(* IEC 61131-3 sources: trust-platform/examples/control/03-production-quality-digital-pid/38-positional-incremental-pid/src, 2 files *)

(* ---- Main.st ---- *)
USING Control;

(* Fraction of the raw-minus-filtered difference applied per update: alpha = dt/(Tf + dt). *)
FUNCTION FilterFraction : LREAL
VAR_INPUT
    CycleTime : LREAL;
    FilterTime : LREAL;
END_VAR
FilterFraction := CycleTime / (FilterTime + CycleTime);
END_FUNCTION

(* One first-order filter update: the filtered value moves alpha of the way toward the raw value. *)
FUNCTION FilterUpdate : LREAL
VAR_INPUT
    PreviousFilteredValue : LREAL;
    RawValue : LREAL;
    FilterFraction : LREAL;
END_VAR
FilterUpdate := PreviousFilteredValue + FilterFraction * (RawValue - PreviousFilteredValue);
END_FUNCTION

FUNCTION SamePidParameters : BOOL
VAR_INPUT
    Left : Control.PIDParameters;
    Right : Control.PIDParameters;
END_VAR
SamePidParameters :=
    Left.ProportionalGain = Right.ProportionalGain
    AND Left.IntegralGain = Right.IntegralGain
    AND Left.DerivativeGain = Right.DerivativeGain
    AND Left.ProportionalSetpointWeight = Right.ProportionalSetpointWeight
    AND Left.DerivativeSetpointWeight = Right.DerivativeSetpointWeight
    AND Left.Bias = Right.Bias
    AND Left.OutputMinimum = Right.OutputMinimum
    AND Left.OutputMaximum = Right.OutputMaximum
    AND Left.RateMinimum = Right.RateMinimum
    AND Left.RateMaximum = Right.RateMaximum
    AND Left.TrackingTime = Right.TrackingTime
    AND Left.AntiWindup = Right.AntiWindup;
END_FUNCTION

(* The positional form of this lesson's PID (β = 1, γ = 0): the complete request every update, from its own
   retained integral. Three rules make it the same controller as the incremental form of Control.PID:
   tracking corrects the integral after the clamp, in Manual the integral follows the manual torque, and a
   gain revision moves the change of the previous P and D into the integral. *)
FUNCTION_BLOCK PositionalPid
VAR_INPUT
    Parameters : Control.PIDParameters;
    Input : Control.PIDInput;
    PreloadOnGainRevision : BOOL := TRUE;
END_VAR
VAR_OUTPUT
    ErrorRad : LREAL;
    ProportionalNm : LREAL;
    TrialIntegralNm : LREAL;
    DerivativeNm : LREAL;
    RequestNm : LREAL;
    TorqueNm : LREAL;
    IntegralNm : LREAL;
END_VAR
VAR
    ProportionalGain : LREAL;
    DerivativeGain : LREAL;
    VelocityRadS : LREAL;
    PreviousAngleRad : LREAL;
    PreviousErrorRad : LREAL;
    PreviousVelocityRadS : LREAL;
END_VAR
(* Gain revision: P and D of the previous update change by (Kp,old − Kp,new)·e and (Kd,new − Kd,old)·ω_f;
   the integral takes that over, so the retained request stays the same. *)
IF PreloadOnGainRevision THEN
    IntegralNm := IntegralNm
        + (ProportionalGain - Parameters.ProportionalGain) * PreviousErrorRad
        - (DerivativeGain - Parameters.DerivativeGain) * PreviousVelocityRadS;
END_IF;
ProportionalGain := Parameters.ProportionalGain;
DerivativeGain := Parameters.DerivativeGain;

ErrorRad := Input.Setpoint - Input.ProcessValue;
VelocityRadS := (Input.ProcessValue - PreviousAngleRad) / Input.CycleTime;
ProportionalNm := ProportionalGain * ErrorRad;
DerivativeNm := -DerivativeGain * VelocityRadS;
IF Input.Mode = PIDMode#Auto THEN
    TrialIntegralNm := IntegralNm + Parameters.IntegralGain * ErrorRad * Input.CycleTime;
    RequestNm := ProportionalNm + TrialIntegralNm + DerivativeNm;
    TorqueNm := LIMIT(Parameters.OutputMinimum, RequestNm, Parameters.OutputMaximum);
    IntegralNm := TrialIntegralNm + Input.CycleTime / Parameters.TrackingTime * (TorqueNm - RequestNm);
ELSE
    (* Manual: the integral follows the manual torque, so the first Auto update continues from it. *)
    RequestNm := Input.ManualOutput;
    TorqueNm := LIMIT(Parameters.OutputMinimum, Input.ManualOutput, Parameters.OutputMaximum);
    IntegralNm := Input.ManualOutput - ProportionalNm - DerivativeNm;
    TrialIntegralNm := IntegralNm;
END_IF;
PreviousAngleRad := Input.ProcessValue;
PreviousErrorRad := ErrorRad;
PreviousVelocityRadS := VelocityRadS;
END_FUNCTION_BLOCK

PROGRAM Main
VAR
    Controller : Control.PID;
    (* The discrete PID of Lesson 38: Kp = 16 N·m/rad, Ki = 4 N·m/(rad·s), Kd = 7 N·m·s/rad on the
       filtered angle, the full target change in P, ±20 N·m with back-calculation (Tt = 1 s). *)
    Parameters : Control.PIDParameters := (
        ProportionalGain := LREAL#16.0,
        IntegralGain := LREAL#4.0,
        DerivativeGain := LREAL#7.0,
        ProportionalSetpointWeight := LREAL#1.0,
        DerivativeSetpointWeight := LREAL#0.0,
        Bias := LREAL#0.0,
        OutputMinimum := LREAL#-20.0,
        OutputMaximum := LREAL#20.0,
        RateMinimum := LREAL#-10000.0,
        RateMaximum := LREAL#10000.0,
        TrackingTime := LREAL#1.0,
        AntiWindup := PIDAntiWindup#BackCalculation
    );
    ConfiguredParameters : Control.PIDParameters;
    ParameterRevision : DINT := 0;
    InitialState : Control.PIDInitialState;
    Input : Control.PIDInput;
    Initialized : BOOL := FALSE;
    AutoMode : BOOL := FALSE;
    ManualTorqueNm : LREAL := 0.0;
    SafetyAbort : BOOL := FALSE;
    SetpointRad : LREAL := 0.0;
    AngleRad : LREAL := 0.0;
    VelocityRadS : LREAL := 0.0;
    TorqueNm : LREAL := 0.0;
    (* Drum load of the simulated test rig, in N·m: the experiment couples a 2 kg weight at the 0.1 m drum
       radius, 1.962 N·m. The controller does not use it. *)
    LoadTorqueNm : LREAL := 0.0;
    (* Measurement filter on the angle: Control.PID differentiates the filtered angle, so D uses the
       filtered velocity. Tf = 0 bypasses the filter. *)
    FilterTimeS : LREAL := 0.1;
    FilterAlpha : LREAL := 1.0;
    FilteredAngleRad : LREAL := 0.0;
    FilterActive : BOOL := FALSE;
    FilterWasActive : BOOL := FALSE;
    (* Three other forms, each updated from the same Input as Controller. None of them drives the axis. *)
    Positional : PositionalPid;
    Unpreloaded : PositionalPid;
    RetainedApplied : Control.PID;
    RetainedAppliedParameters : Control.PIDParameters;
    PositionalTorqueNm : LREAL := 0.0;
    UnpreloadedTorqueNm : LREAL := 0.0;
    RetainedAppliedTorqueNm : LREAL := 0.0;
    ErrorRad : LREAL := 0.0;
    ProportionalNm : LREAL := 0.0;
    DerivativeNm : LREAL := 0.0;
    RequestNm : LREAL := 0.0;
    IntegralNm : LREAL := 0.0;
    (* Project experiment. *)
    ExperimentEnabled : BOOL := FALSE;
    ExperimentWasEnabled : BOOL := FALSE;
    Active : BOOL := FALSE;
    ExperimentUpdates : DINT := 0;
    GainBeforeRevision : LREAL := 16.0;
    (* Software travel and speed limits of the axis. *)
    AngleLimitRad : LREAL := 2.0;
    VelocityLimitRadS : LREAL := 10.0;
END_VAR

(* Leaving the travel or speed range removes the torque until a full restart. *)
IF ABS(AngleRad) > AngleLimitRad OR ABS(VelocityRadS) > VelocityLimitRadS THEN
    SafetyAbort := TRUE;
END_IF;

(* Control Studio's project experiment couples the drum load and steps the target to 1.5 rad in Auto; 1 s
   later it applies Kp = 24 N·m/rad, as a gain revision would. Its end uncouples the load, restores the gain
   and returns to Manual with zero torque. *)
IF ExperimentEnabled AND NOT ExperimentWasEnabled THEN
    Active := TRUE;
    ExperimentUpdates := 0;
    LoadTorqueNm := LREAL#1.962;
    SetpointRad := LREAL#1.5;
    AutoMode := TRUE;
ELSIF NOT ExperimentEnabled AND ExperimentWasEnabled THEN
    Active := FALSE;
    LoadTorqueNm := LREAL#0.0;
    AutoMode := FALSE;
    SetpointRad := AngleRad;
    IF ExperimentUpdates > 50 THEN
        Parameters.ProportionalGain := GainBeforeRevision;
    END_IF;
END_IF;
ExperimentWasEnabled := ExperimentEnabled;
IF Active THEN
    IF ExperimentUpdates = 50 THEN
        GainBeforeRevision := Parameters.ProportionalGain;
        Parameters.ProportionalGain := LREAL#24.0;
    END_IF;
    ExperimentUpdates := ExperimentUpdates + 1;
END_IF;

(* Control Studio's Apply replaces this complete record at the task boundary. *)
IF NOT Initialized OR NOT SamePidParameters(Left := Parameters, Right := ConfiguredParameters) THEN
    ConfiguredParameters := Parameters;
    ParameterRevision := ParameterRevision + 1;
END_IF;
Controller.Configure(Parameters := Parameters);
(* Tracking with Tt = Δt removes the whole excess: this controller retains the applied torque. *)
RetainedAppliedParameters := Parameters;
RetainedAppliedParameters.TrackingTime := LREAL#0.02;
RetainedApplied.Configure(Parameters := RetainedAppliedParameters);

IF NOT Initialized THEN
    (* Hot reset: the axis rests without torque and the setpoint follows the measured angle. *)
    ManualTorqueNm := LREAL#0.0;
    IF NOT AutoMode THEN
        SetpointRad := AngleRad;
    END_IF;
    InitialState.Setpoint := SetpointRad;
    InitialState.ProcessValue := AngleRad;
    InitialState.NominalOutput := ManualTorqueNm;
    InitialState.SaturatedOutput := ManualTorqueNm;
    InitialState.SetpointRate := LREAL#0.0;
    InitialState.ProcessValueRate := LREAL#0.0;
    InitialState.FeedForward := LREAL#0.0;
    Controller.Initialize(State := InitialState);
    RetainedApplied.Initialize(State := InitialState);
    Initialized := TRUE;
END_IF;

(* The filter runs while the controller is in Auto. In Manual and in the Auto-entry scan it restarts
   from the measurement, so entering Auto is exactly bumpless; filtering starts with the next scan. *)
FilterAlpha := FilterFraction(CycleTime := LREAL#0.02, FilterTime := MAX(FilterTimeS, LREAL#0.0));
FilterActive := AutoMode AND NOT SafetyAbort AND Parameters.ProportionalGain > LREAL#0.0;
IF FilterActive AND FilterWasActive THEN
    FilteredAngleRad := FilterUpdate(PreviousFilteredValue := FilteredAngleRad, RawValue := AngleRad, FilterFraction := FilterAlpha);
ELSE
    FilteredAngleRad := AngleRad;
END_IF;
FilterWasActive := FilterActive;

Input.Setpoint := SetpointRad;
Input.ProcessValue := FilteredAngleRad;
Input.CycleTime := LREAL#0.02;
Input.FeedForward := LREAL#0.0;
Input.TrackingOutput := ManualTorqueNm;
IF SafetyAbort THEN
    Input.Mode := PIDMode#Manual;
    Input.ManualOutput := LREAL#0.0;
ELSIF AutoMode AND Parameters.ProportionalGain > LREAL#0.0 THEN
    Input.Mode := PIDMode#Auto;
    Input.ManualOutput := ManualTorqueNm;
ELSE
    Input.Mode := PIDMode#Manual;
    Input.ManualOutput := ManualTorqueNm;
END_IF;
TorqueNm := Controller.Update(Input := Input);

(* The positional form with its three rules, the same form without the gain-revision rule, and Control.PID
   retaining the applied torque. *)
Positional(Parameters := Parameters, Input := Input);
Unpreloaded(Parameters := Parameters, Input := Input, PreloadOnGainRevision := FALSE);
RetainedAppliedTorqueNm := RetainedApplied.Update(Input := Input);
PositionalTorqueNm := Positional.TorqueNm;
UnpreloadedTorqueNm := Unpreloaded.TorqueNm;
ErrorRad := Positional.ErrorRad;
ProportionalNm := Positional.ProportionalNm;
DerivativeNm := Positional.DerivativeNm;
RequestNm := Positional.RequestNm;
IntegralNm := Positional.IntegralNm;

END_PROGRAM

CONFIGURATION Config
RESOURCE Res ON PLC
    TASK MainTask(INTERVAL := T#20ms, PRIORITY := 1);
    PROGRAM P1 WITH MainTask : Main;
END_RESOURCE
VAR_CONFIG
    P1.SafetyAbort AT %MX24.0 : BOOL;
    P1.TorqueNm AT %QL0 : LREAL;
    P1.LoadTorqueNm AT %QL8 : LREAL;
    P1.AngleRad AT %IL0 : LREAL;
    P1.VelocityRadS AT %IL8 : LREAL;
    P1.SetpointRad AT %ML0 : LREAL;
    P1.ManualTorqueNm AT %ML8 : LREAL;
    P1.FilteredAngleRad AT %ML32 : LREAL;
    P1.ErrorRad AT %ML40 : LREAL;
    P1.ProportionalNm AT %ML48 : LREAL;
    P1.DerivativeNm AT %ML64 : LREAL;
    P1.RequestNm AT %ML72 : LREAL;
    P1.IntegralNm AT %ML80 : LREAL;
    P1.ExperimentEnabled AT %MX88.0 : BOOL;
    P1.Active AT %MX88.1 : BOOL;
    P1.PositionalTorqueNm AT %ML96 : LREAL;
    P1.RetainedAppliedTorqueNm AT %ML104 : LREAL;
    P1.UnpreloadedTorqueNm AT %ML112 : LREAL;
END_VAR
END_CONFIGURATION

(* ---- tests.st ---- *)
(* @trustlsp:runtime-ignore — run these assertions with trust-dev test;
   they are not scheduled PLC instances in the lesson simulator. *)
USING Control;

TEST_PROGRAM TheIncrementOfTheExample
VAR
    Increment : LREAL;
    Controller : Control.PID;
    Parameters : Control.PIDParameters;
    State : Control.PIDInitialState;
    Input : Control.PIDInput;
END_VAR
(* e 0.10 → 0.096 rad, ω_f 0.20 → 0.22 rad/s, Kp 16, Ki 4, Kd 7, Δt 0.02 s, no tracking correction. *)
Increment := LREAL#16.0 * (LREAL#0.096 - LREAL#0.10) + LREAL#4.0 * LREAL#0.096 * LREAL#0.02
    - LREAL#7.0 * (LREAL#0.22 - LREAL#0.20);
ASSERT_NEAR(EXPECTED := LREAL#-0.19632, ACTUAL := Increment, DELTA := LREAL#1.0e-12);
ASSERT_NEAR(EXPECTED := LREAL#1.00368, ACTUAL := LREAL#1.2 + Increment, DELTA := LREAL#1.0e-12);
(* Control.PID adds the same increment to its retained 1.2 N·m. The angle moves 0.004 rad and then 0.0044 rad
   per update (0.20 and 0.22 rad/s) while the target moves 0.0004 rad: the error goes from 0.10 to 0.096 rad. *)
Parameters.ProportionalGain := LREAL#16.0;
Parameters.IntegralGain := LREAL#4.0;
Parameters.DerivativeGain := LREAL#7.0;
Parameters.ProportionalSetpointWeight := LREAL#1.0;
Parameters.OutputMinimum := LREAL#-20.0;
Parameters.OutputMaximum := LREAL#20.0;
Parameters.RateMinimum := LREAL#-10000.0;
Parameters.RateMaximum := LREAL#10000.0;
Parameters.TrackingTime := LREAL#1.0;
Parameters.AntiWindup := PIDAntiWindup#BackCalculation;
Controller.Configure(Parameters := Parameters);
State.Setpoint := LREAL#0.5;
State.ProcessValue := LREAL#0.4;
State.ProcessValueRate := LREAL#0.20;
State.NominalOutput := LREAL#1.2;
State.SaturatedOutput := LREAL#1.2;
Controller.Initialize(State := State);
Input.Mode := PIDMode#Auto;
Input.CycleTime := LREAL#0.02;
Input.Setpoint := LREAL#0.5004;
Input.ProcessValue := LREAL#0.4044;
ASSERT_NEAR(EXPECTED := LREAL#1.00368, ACTUAL := Controller.Update(Input := Input), DELTA := LREAL#1.0e-9);
END_TEST_PROGRAM

TEST_PROGRAM TheClampedUpdateRetainsTheCorrectedRequest
VAR
    Controller : Control.PID;
    RetainedApplied : Control.PID;
    Parameters : Control.PIDParameters;
    State : Control.PIDInitialState;
    Input : Control.PIDInput;
END_VAR
(* The previous update requested 25 N·m against the 20 N·m limit. At rest on target the increment is zero, so
   this update requests 25 N·m again and the drive gets 20 N·m. *)
Parameters.ProportionalGain := LREAL#16.0;
Parameters.IntegralGain := LREAL#4.0;
Parameters.DerivativeGain := LREAL#7.0;
Parameters.ProportionalSetpointWeight := LREAL#1.0;
Parameters.OutputMinimum := LREAL#-20.0;
Parameters.OutputMaximum := LREAL#20.0;
Parameters.RateMinimum := LREAL#-10000.0;
Parameters.RateMaximum := LREAL#10000.0;
Parameters.TrackingTime := LREAL#1.0;
Parameters.AntiWindup := PIDAntiWindup#BackCalculation;
Controller.Configure(Parameters := Parameters);
State.Setpoint := LREAL#0.5;
State.ProcessValue := LREAL#0.5;
State.NominalOutput := LREAL#25.0;
State.SaturatedOutput := LREAL#20.0;
Controller.Initialize(State := State);
Input.Mode := PIDMode#Auto;
Input.CycleTime := LREAL#0.02;
Input.Setpoint := LREAL#0.5;
Input.ProcessValue := LREAL#0.5;
ASSERT_NEAR(EXPECTED := LREAL#20.0, ACTUAL := Controller.Update(Input := Input), DELTA := LREAL#1.0e-12);
(* γ = (Δt/Tt)(u_a − u_r) = 0.02 · (20 − 25) = −0.1 N·m: the retained request is 24.9 N·m. *)
State := Controller.GetState();
ASSERT_NEAR(EXPECTED := LREAL#24.9, ACTUAL := State.NominalOutput, DELTA := LREAL#1.0e-9);
(* Tracking with Tt = Δt removes the whole excess: that controller retains the applied 20 N·m. *)
Parameters.TrackingTime := LREAL#0.02;
RetainedApplied.Configure(Parameters := Parameters);
State.NominalOutput := LREAL#25.0;
State.SaturatedOutput := LREAL#20.0;
RetainedApplied.Initialize(State := State);
ASSERT_NEAR(EXPECTED := LREAL#20.0, ACTUAL := RetainedApplied.Update(Input := Input), DELTA := LREAL#1.0e-12);
State := RetainedApplied.GetState();
ASSERT_NEAR(EXPECTED := LREAL#20.0, ACTUAL := State.NominalOutput, DELTA := LREAL#1.0e-12);
END_TEST_PROGRAM

TEST_PROGRAM AGainRevisionAtConstantError
VAR
    Controller : Control.PID;
    Positional : PositionalPid;
    Unpreloaded : PositionalPid;
    Parameters : Control.PIDParameters;
    State : Control.PIDInitialState;
    Input : Control.PIDInput;
    Count : INT;
    Before : LREAL;
    After : LREAL;
END_VAR
(* The axis rests 0.1 rad below its target. Two Manual updates hold 1.6 N·m; then one Auto update with
   Kp = 16, and one after the revision to Kp = 24. *)
Parameters.ProportionalGain := LREAL#16.0;
Parameters.IntegralGain := LREAL#4.0;
Parameters.DerivativeGain := LREAL#7.0;
Parameters.ProportionalSetpointWeight := LREAL#1.0;
Parameters.OutputMinimum := LREAL#-20.0;
Parameters.OutputMaximum := LREAL#20.0;
Parameters.RateMinimum := LREAL#-10000.0;
Parameters.RateMaximum := LREAL#10000.0;
Parameters.TrackingTime := LREAL#1.0;
Parameters.AntiWindup := PIDAntiWindup#BackCalculation;
Controller.Configure(Parameters := Parameters);
State.Setpoint := LREAL#0.5;
State.ProcessValue := LREAL#0.4;
Controller.Initialize(State := State);
Input.CycleTime := LREAL#0.02;
Input.Setpoint := LREAL#0.5;
Input.ProcessValue := LREAL#0.4;
Input.ManualOutput := LREAL#1.6;
Input.Mode := PIDMode#Manual;
FOR Count := 1 TO 2 DO
    Controller.Update(Input := Input);
    Positional(Parameters := Parameters, Input := Input);
    Unpreloaded(Parameters := Parameters, Input := Input, PreloadOnGainRevision := FALSE);
END_FOR;
Input.Mode := PIDMode#Auto;
Before := Controller.Update(Input := Input);
Positional(Parameters := Parameters, Input := Input);
Unpreloaded(Parameters := Parameters, Input := Input, PreloadOnGainRevision := FALSE);
(* 1.6 + Ki·e·Δt = 1.6 + 4 · 0.1 · 0.02 = 1.608 N·m in both forms. *)
ASSERT_NEAR(EXPECTED := LREAL#1.608, ACTUAL := Before, DELTA := LREAL#1.0e-12);
ASSERT_NEAR(EXPECTED := Before, ACTUAL := Positional.TorqueNm, DELTA := LREAL#1.0e-12);
Parameters.ProportionalGain := LREAL#24.0;
Controller.Configure(Parameters := Parameters);
After := Controller.Update(Input := Input);
Positional(Parameters := Parameters, Input := Input);
Unpreloaded(Parameters := Parameters, Input := Input, PreloadOnGainRevision := FALSE);
(* The error did not change, so Control.PID adds only the integral increment. *)
ASSERT_NEAR(EXPECTED := LREAL#1.616, ACTUAL := After, DELTA := LREAL#1.0e-12);
(* P rises by (24 − 16) · 0.1 = 0.8 N·m; the preloaded integral takes it over, so the positional torque agrees. *)
ASSERT_NEAR(EXPECTED := LREAL#2.4, ACTUAL := Positional.ProportionalNm, DELTA := LREAL#1.0e-12);
ASSERT_NEAR(EXPECTED := After, ACTUAL := Positional.TorqueNm, DELTA := LREAL#1.0e-12);
(* Without the preload the positional torque jumps by 0.8 N·m. *)
ASSERT_NEAR(EXPECTED := After + LREAL#0.8, ACTUAL := Unpreloaded.TorqueNm, DELTA := LREAL#1.0e-12);
END_TEST_PROGRAM
